TYPE ST_Recipe :
STRUCT
	sName		: STRING(31);
	fTargetLevel	: T_Percent := 80;
	tSettle		: TIME := T#2S;
END_STRUCT
END_TYPE

(* stored: Version 1.1.0.1
   DUT ST_Recipe: Id {4a4f9780-4f3b-4d61-8087-108410ca57d2} *)
